  movel([-0.151447, -0.814996, -2.788348, -1.109046, 1.570796, 1.419350],accel_mss,speed_ms,0,blend_radius_m)
  movel([-0.155435, -0.823121, -2.786879, -1.102389, 1.570796, 1.415362],accel_mss,speed_ms,0,blend_radius_m)
  movel([-0.157149, -0.827095, -2.786148, -1.099146, 1.570796, 1.413648],accel_mss,speed_ms,0,blend_radius_m)
  movel([-0.159989, -0.834849, -2.784696, -1.092844, 1.570796, 1.410807],accel_mss,speed_ms,0,blend_radius_m)
  movel([-0.161109, -0.838634, -2.783975, -1.089780, 1.570796, 1.409688],accel_mss,speed_ms,0,blend_radius_m)
  movel([-0.162732, -0.846011, -2.782547, -1.083831, 1.570796, 1.408064],accel_mss,speed_ms,0,blend_radius_m)
  movel([-0.163230, -0.849609, -2.781839, -1.080941, 1.570796, 1.407566],accel_mss,speed_ms,0,blend_radius_m)
  movel([-0.163513, -0.853139, -2.781138, -1.078112, 1.570796, 1.407283],accel_mss,speed_ms,0,blend_radius_m)
  movel([-0.163602, -0.858015, -2.780157, -1.074217, 1.570796, 1.407194],accel_mss,speed_ms,0,blend_radius_m)
  movel([-0.163380, -0.862704, -2.779201, -1.070483, 1.570796, 1.407417],accel_mss,speed_ms,0,blend_radius_m)
  movel([-0.162870, -0.867194, -2.778274, -1.066921, 1.570796, 1.407926],accel_mss,speed_ms,0,blend_radius_m)
  movel([-0.162104, -0.871488, -2.777376, -1.063525, 1.570796, 1.408692],accel_mss,speed_ms,0,blend_radius_m)
  movel([-0.161097, -0.875560, -2.776515, -1.060315, 1.570796, 1.409700],accel_mss,speed_ms,0,blend_radius_m)
  movel([-0.159870, -0.879398, -2.775693, -1.057297, 1.570796, 1.410927],accel_mss,speed_ms,0,blend_radius_m)
  movel([-0.158448, -0.882999, -2.774915, -1.054475, 1.570796, 1.412348],accel_mss,speed_ms,0,blend_radius_m)
  movel([-0.156848, -0.886344, -2.774185, -1.051861, 1.570796, 1.413948],accel_mss,speed_ms,0,blend_radius_m)
  movel([-0.149158, -0.898055, -2.771574, -1.042759, 1.570796, 1.421638],accel_mss,speed_ms,0,blend_radius_m)
  movel([-0.143209, -0.907609, -2.769382, -1.035398, 1.570796, 1.427587],accel_mss,speed_ms,0,blend_radius_m)
  movel([-0.142775, -0.908633, -2.769143, -1.034613, 1.570796, 1.428021],accel_mss,speed_ms,0,blend_radius_m)
  movel([-0.135600, -0.899262, -2.771300, -1.041826, 1.570796, 1.435197],accel_mss,speed_ms,0,blend_radius_m)
  movel([-0.127938, -0.890014, -2.773376, -1.048999, 1.570796, 1.442859],accel_mss,speed_ms,0,blend_radius_m)
  movel([-0.119839, -0.880922, -2.775365, -1.056102, 1.570796, 1.450957],accel_mss,speed_ms,0,blend_radius_m)
  movel([-0.111369, -0.872030, -2.777262, -1.063097, 1.570796, 1.459427],accel_mss,speed_ms,0,blend_radius_m)
  movel([-0.102591, -0.863390, -2.779061, -1.069938, 1.570796, 1.468205],accel_mss,speed_ms,0,blend_radius_m)
  movel([-0.093574, -0.855040, -2.780757, -1.076592, 1.570796, 1.477222],accel_mss,speed_ms,0,blend_radius_m)
  movel([-0.084386, -0.847036, -2.782346, -1.083007, 1.570796, 1.486410],accel_mss,speed_ms,0,blend_radius_m)
  movel([-0.075105, -0.839424, -2.783823, -1.089142, 1.570796, 1.495692],accel_mss,speed_ms,0,blend_radius_m)
  movel([-0.070692, -0.836034, -2.784471, -1.091884, 1.570796, 1.500104],accel_mss,speed_ms,0,blend_radius_m)
  movel([-0.066171, -0.832804, -2.785082, -1.094503, 1.570796, 1.504626],accel_mss,speed_ms,0,blend_radius_m)
  movel([-0.061579, -0.829772, -2.785650, -1.096967, 1.570796, 1.509218],accel_mss,speed_ms,0,blend_radius_m)
  movel([-0.056967, -0.826981, -2.786169, -1.099239, 1.570796, 1.513830],accel_mss,speed_ms,0,blend_radius_m)
  movel([-0.052375, -0.824471, -2.786631, -1.101286, 1.570796, 1.518421],accel_mss,speed_ms,0,blend_radius_m)
  movel([-0.047846, -0.822284, -2.787032, -1.103074, 1.570796, 1.522951],accel_mss,speed_ms,0,blend_radius_m)
  movel([-0.043425, -0.820455, -2.787365, -1.104569, 1.570796, 1.527371],accel_mss,speed_ms,0,blend_radius_m)
  movel([-0.039161, -0.819026, -2.787624, -1.105740, 1.570796, 1.531636],accel_mss,speed_ms,0,blend_radius_m)
  movel([-0.035094, -0.818037, -2.787802, -1.106550, 1.570796, 1.535702],accel_mss,speed_ms,0,blend_radius_m)
  movel([-0.031268, -0.817523, -2.787894, -1.106971, 1.570796, 1.539528],accel_mss,speed_ms,0,blend_radius_m)
  movel([-0.027734, -0.817526, -2.787894, -1.106969, 1.570796, 1.543062],accel_mss,speed_ms,0,blend_radius_m)
  movel([-0.024533, -0.818078, -2.787795, -1.106516, 1.570796, 1.546264],accel_mss,speed_ms,0,blend_radius_m)
  movel([-0.021709, -0.819214, -2.787590, -1.105586, 1.570796, 1.549087],accel_mss,speed_ms,0,blend_radius_m)
  movel([-0.019297, -0.820962, -2.787273, -1.104155, 1.570796, 1.551499],accel_mss,speed_ms,0,blend_radius_m)
  movel([-0.017345, -0.823352, -2.786837, -1.102201, 1.570796, 1.553452],accel_mss,speed_ms,0,blend_radius_m)
  movel([-0.015891, -0.826416, -2.786273, -1.099700, 1.570796, 1.554905],accel_mss,speed_ms,0,blend_radius_m)
  movel([-0.014708, -0.831178, -2.785387, -1.095824, 1.570796, 1.556088],accel_mss,speed_ms,0,blend_radius_m)
  movel([-0.014174, -0.836590, -2.784365, -1.091434, 1.570796, 1.556622],accel_mss,speed_ms,0,blend_radius_m)
  movel([-0.014196, -0.842501, -2.783230, -1.086658, 1.570796, 1.556600],accel_mss,speed_ms,0,blend_radius_m)
  movel([-0.014673, -0.848767, -2.782005, -1.081616, 1.570796, 1.556123],accel_mss,speed_ms,0,blend_radius_m)
  movel([-0.015515, -0.855244, -2.780716, -1.076429, 1.570796, 1.555282],accel_mss,speed_ms,0,blend_radius_m)
  movel([-0.016634, -0.861800, -2.779387, -1.071202, 1.570796, 1.554162],accel_mss,speed_ms,0,blend_radius_m)
  movel([-0.019330, -0.874610, -2.776716, -1.061062, 1.570796, 1.551466],accel_mss,speed_ms,0,blend_radius_m)
  movel([-0.021385, -0.882738, -2.774972, -1.054680, 1.570796, 1.549411],accel_mss,speed_ms,0,blend_radius_m)
  movel([-0.023782, -0.890821, -2.773197, -1.048372, 1.570796, 1.547015],accel_mss,speed_ms,0,blend_radius_m)
  movel([-0.026474, -0.898860, -2.771392, -1.042138, 1.570796, 1.544323],accel_mss,speed_ms,0,blend_radius_m)
  movel([-0.029419, -0.906874, -2.769553, -1.035963, 1.570796, 1.541377],accel_mss,speed_ms,0,blend_radius_m)
  movel([-0.032573, -0.914860, -2.767679, -1.029850, 1.570796, 1.538223],accel_mss,speed_ms,0,blend_radius_m)
  movel([-0.035892, -0.922833, -2.765768, -1.023788, 1.570796, 1.534904],accel_mss,speed_ms,0,blend_radius_m)
  movel([-0.042880, -0.938782, -2.761820, -1.011787, 1.570796, 1.527916],accel_mss,speed_ms,0,blend_radius_m)
  movel([-0.036325, -0.939075, -2.761746, -1.011568, 1.570796, 1.534471],accel_mss,speed_ms,0,blend_radius_m)
  movel([-0.032953, -0.939481, -2.761643, -1.011265, 1.570796, 1.537843],accel_mss,speed_ms,0,blend_radius_m)
  movel([-0.030089, -0.940387, -2.761414, -1.010589, 1.570796, 1.540707],accel_mss,speed_ms,0,blend_radius_m)
  movel([-0.028984, -0.941104, -2.761231, -1.010053, 1.570796, 1.541813],accel_mss,speed_ms,0,blend_radius_m)
  movel([-0.028168, -0.942040, -2.760993, -1.009356, 1.570796, 1.542628],accel_mss,speed_ms,0,blend_radius_m)
  movel([-0.027690, -0.943217, -2.760692, -1.008479, 1.570796, 1.543106],accel_mss,speed_ms,0,blend_radius_m)
  movel([-0.027603, -0.944666, -2.760321, -1.007402, 1.570796, 1.543193],accel_mss,speed_ms,0,blend_radius_m)
  movel([-0.027958, -0.946409, -2.759872, -1.006107, 1.570796, 1.542838],accel_mss,speed_ms,0,blend_radius_m)
  movel([-0.028810, -0.948485, -2.759335, -1.004569, 1.570796, 1.541986],accel_mss,speed_ms,0,blend_radius_m)
  movel([-0.030204, -0.950916, -2.758703, -1.002770, 1.570796, 1.540592],accel_mss,speed_ms,0,blend_radius_m)
  movel([-0.032189, -0.953722, -2.757967, -1.000700, 1.570796, 1.538607],accel_mss,speed_ms,0,blend_radius_m)
  movel([-0.034030, -0.956006, -2.757365, -0.999018, 1.570796, 1.536766],accel_mss,speed_ms,0,blend_radius_m)
  movel([-0.035882, -0.958061, -2.756820, -0.997508, 1.570796, 1.534914],accel_mss,speed_ms,0,blend_radius_m)
  movel([-0.037742, -0.959903, -2.756328, -0.996157, 1.570796, 1.533055],accel_mss,speed_ms,0,blend_radius_m)
  movel([-0.041487, -0.963031, -2.755489, -0.993869, 1.570796, 1.529310],accel_mss,speed_ms,0,blend_radius_m)
  movel([-0.043369, -0.964351, -2.755133, -0.992905, 1.570796, 1.527427],accel_mss,speed_ms,0,blend_radius_m)
  movel([-0.047159, -0.966604, -2.754522, -0.991264, 1.570796, 1.523638],accel_mss,speed_ms,0,blend_radius_m)
  movel([-0.050963, -0.968447, -2.754019, -0.989923, 1.570796, 1.519833],accel_mss,speed_ms,0,blend_radius_m)
  movel([-0.054779, -0.970023, -2.753588, -0.988778, 1.570796, 1.516017],accel_mss,speed_ms,0,blend_radius_m)
  movel([-0.062394, -0.972906, -2.752793, -0.986690, 1.570796, 1.508402],accel_mss,speed_ms,0,blend_radius_m)
  movel([-0.066370, -0.979281, -2.751016, -0.982092, 1.570796, 1.504426],accel_mss,speed_ms,0,blend_radius_m)
  movel([-0.068546, -0.982465, -2.750118, -0.979807, 1.570796, 1.502250],accel_mss,speed_ms,0,blend_radius_m)
  movel([-0.070857, -0.985559, -2.749237, -0.977593, 1.570796, 1.499939],accel_mss,speed_ms,0,blend_radius_m)
  movel([-0.073309, -0.988496, -2.748395, -0.975498, 1.570796, 1.497488],accel_mss,speed_ms,0,blend_radius_m)
  movel([-0.075903, -0.991209, -2.747612, -0.973569, 1.570796, 1.494894],accel_mss,speed_ms,0,blend_radius_m)
  movel([-0.078648, -0.993632, -2.746907, -0.971850, 1.570796, 1.492149],accel_mss,speed_ms,0,blend_radius_m)
  movel([-0.081555, -0.995707, -2.746300, -0.970382, 1.570796, 1.489241],accel_mss,speed_ms,0,blend_radius_m)
  movel([-0.083598, -0.996753, -2.745993, -0.969643, 1.570796, 1.487198],accel_mss,speed_ms,0,blend_radius_m)
  movel([-0.085214, -0.997109, -2.745888, -0.969392, 1.570796, 1.485582],accel_mss,speed_ms,0,blend_radius_m)
  movel([-0.086450, -0.996877, -2.745957, -0.969556, 1.570796, 1.484347],accel_mss,speed_ms,0,blend_radius_m)
  movel([-0.087346, -0.996152, -2.746170, -0.970067, 1.570796, 1.483451],accel_mss,speed_ms,0,blend_radius_m)
  movel([-0.087946, -0.995031, -2.746498, -0.970860, 1.570796, 1.482851],accel_mss,speed_ms,0,blend_radius_m)
  movel([-0.088287, -0.993617, -2.746911, -0.971861, 1.570796, 1.482509],accel_mss,speed_ms,0,blend_radius_m)
  movel([-0.088418, -0.992006, -2.747380, -0.973003, 1.570796, 1.482378],accel_mss,speed_ms,0,blend_radius_m)
  movel([-0.088369, -0.990291, -2.747877, -0.974221, 1.570796, 1.482428],accel_mss,speed_ms,0,blend_radius_m)
  movel([-0.087893, -0.986486, -2.748972, -0.976931, 1.570796, 1.482904],accel_mss,speed_ms,0,blend_radius_m)
  movel([-0.087059, -0.982547, -2.750094, -0.979748, 1.570796, 1.483737],accel_mss,speed_ms,0,blend_radius_m)
  movel([-0.084858, -0.974333, -2.752398, -0.985658, 1.570796, 1.485939],accel_mss,speed_ms,0,blend_radius_m)
  movel([-0.093540, -0.972916, -2.752791, -0.986682, 1.570796, 1.477256],accel_mss,speed_ms,0,blend_radius_m)
  movel([-0.102455, -0.971877, -2.753077, -0.987434, 1.570796, 1.468341],accel_mss,speed_ms,0,blend_radius_m)
  movel([-0.111365, -0.970808, -2.753372, -0.988209, 1.570796, 1.459431],accel_mss,speed_ms,0,blend_radius_m)
  movel([-0.115747, -0.970134, -2.753557, -0.988698, 1.570796, 1.455049],accel_mss,speed_ms,0,blend_radius_m)
  movel([-0.120046, -0.969296, -2.753787, -0.989306, 1.570796, 1.450750],accel_mss,speed_ms,0,blend_radius_m)
  movel([-0.124039, -0.968285, -2.754064, -0.990041, 1.570796, 1.446757],accel_mss,speed_ms,0,blend_radius_m)
  movel([-0.127889, -0.967094, -2.754388, -0.990906, 1.570796, 1.442907],accel_mss,speed_ms,0,blend_radius_m)
  movel([-0.135327, -0.964371, -2.755127, -0.992891, 1.570796, 1.435469],accel_mss,speed_ms,0,blend_radius_m)
  movel([-0.142709, -0.961582, -2.755879, -0.994928, 1.570796, 1.428087],accel_mss,speed_ms,0,blend_radius_m)
  movel([-0.150371, -0.959179, -2.756522, -0.996688, 1.570796, 1.420425],accel_mss,speed_ms,0,blend_radius_m)
  movel([-0.152086, -0.963930, -2.755246, -0.993213, 1.570796, 1.418710],accel_mss,speed_ms,0,blend_radius_m)
  movel([-0.153549, -0.968557, -2.753989, -0.989843, 1.570796, 1.417247],accel_mss,speed_ms,0,blend_radius_m)
  movel([-0.154762, -0.973052, -2.752753, -0.986584, 1.570796, 1.416035],accel_mss,speed_ms,0,blend_radius_m)
  movel([-0.155729, -0.977408, -2.751541, -0.983440, 1.570796, 1.415067],accel_mss,speed_ms,0,blend_radius_m)
  movel([-0.156451, -0.981621, -2.750356, -0.980411, 1.570796, 1.414345],accel_mss,speed_ms,0,blend_radius_m)
  movel([-0.156938, -0.985687, -2.749200, -0.977501, 1.570796, 1.413859],accel_mss,speed_ms,0,blend_radius_m)
  movel([-0.157185, -0.989600, -2.748077, -0.974712, 1.570796, 1.413612],accel_mss,speed_ms,0,blend_radius_m)
  movel([-0.157205, -0.993359, -2.746986, -0.972043, 1.570796, 1.413592],accel_mss,speed_ms,0,blend_radius_m)
  movel([-0.156995, -0.996957, -2.745933, -0.969499, 1.570796, 1.413802],accel_mss,speed_ms,0,blend_radius_m)
  movel([-0.156554, -1.000385, -2.744920, -0.967083, 1.570796, 1.414242],accel_mss,speed_ms,0,blend_radius_m)
  movel([-0.155895, -1.003650, -2.743948, -0.964791, 1.570796, 1.414901],accel_mss,speed_ms,0,blend_radius_m)
  movel([-0.155018, -1.006740, -2.743020, -0.962629, 1.570796, 1.415778],accel_mss,speed_ms,0,blend_radius_m)
  movel([-0.153919, -1.009647, -2.742140, -0.960602, 1.570796, 1.416877],accel_mss,speed_ms,0,blend_radius_m)
  movel([-0.152607, -1.012377, -2.741308, -0.958704, 1.570796, 1.418189],accel_mss,speed_ms,0,blend_radius_m)
  movel([-0.151084, -1.014919, -2.740528, -0.956942, 1.570796, 1.419713],accel_mss,speed_ms,0,blend_radius_m)
  movel([-0.149346, -1.017271, -2.739802, -0.955317, 1.570796, 1.421450],accel_mss,speed_ms,0,blend_radius_m)
  movel([-0.146282, -1.020526, -2.738789, -0.953073, 1.570796, 1.424514],accel_mss,speed_ms,0,blend_radius_m)
  movel([-0.142850, -1.023308, -2.737918, -0.951163, 1.570796, 1.427946],accel_mss,speed_ms,0,blend_radius_m)
  movel([-0.139097, -1.025667, -2.737174, -0.949548, 1.570796, 1.431699],accel_mss,speed_ms,0,blend_radius_m)
  movel([-0.135055, -1.027644, -2.736547, -0.948198, 1.570796, 1.435741],accel_mss,speed_ms,0,blend_radius_m)
  movel([-0.130770, -1.029287, -2.736024, -0.947078, 1.570796, 1.440026],accel_mss,speed_ms,0,blend_radius_m)
  movel([-0.126280, -1.030634, -2.735593, -0.946162, 1.570796, 1.444516],accel_mss,speed_ms,0,blend_radius_m)
  movel([-0.121626, -1.031732, -2.735241, -0.945416, 1.570796, 1.449171],accel_mss,speed_ms,0,blend_radius_m)
  movel([-0.116838, -1.032609, -2.734959, -0.944821, 1.570796, 1.453958],accel_mss,speed_ms,0,blend_radius_m)
  movel([-0.106974, -1.033936, -2.734531, -0.943921, 1.570796, 1.463822],accel_mss,speed_ms,0,blend_radius_m)
  movel([-0.096981, -1.035022, -2.734180, -0.943187, 1.570796, 1.473815],accel_mss,speed_ms,0,blend_radius_m)
  movel([-0.089406, -1.036121, -2.733824, -0.942444, 1.570796, 1.481391],accel_mss,speed_ms,0,blend_radius_m)
  movel([-0.086797, -1.036293, -2.733768, -0.942328, 1.570796, 1.484000],accel_mss,speed_ms,0,blend_radius_m)
  movel([-0.082087, -1.036201, -2.733798, -0.942390, 1.570796, 1.488709],accel_mss,speed_ms,0,blend_radius_m)
  movel([-0.081105, -1.036377, -2.733741, -0.942271, 1.570796, 1.489692],accel_mss,speed_ms,0,blend_radius_m)
  movel([-0.080223, -1.036750, -2.733620, -0.942019, 1.570796, 1.490574],accel_mss,speed_ms,0,blend_radius_m)
  movel([-0.079458, -1.037384, -2.733413, -0.941592, 1.570796, 1.491338],accel_mss,speed_ms,0,blend_radius_m)
  movel([-0.078830, -1.038339, -2.733102, -0.940948, 1.570796, 1.491966],accel_mss,speed_ms,0,blend_radius_m)
  movel([-0.078371, -1.039682, -2.732663, -0.940044, 1.570796, 1.492426],accel_mss,speed_ms,0,blend_radius_m)
  movel([-0.078211, -1.041203, -2.732164, -0.939022, 1.570796, 1.492585],accel_mss,speed_ms,0,blend_radius_m)
  movel([-0.078322, -1.042870, -2.731615, -0.937905, 1.570796, 1.492474],accel_mss,speed_ms,0,blend_radius_m)
  movel([-0.078680, -1.044666, -2.731020, -0.936703, 1.570796, 1.492116],accel_mss,speed_ms,0,blend_radius_m)
  movel([-0.079260, -1.046558, -2.730392, -0.935440, 1.570796, 1.491536],accel_mss,speed_ms,0,blend_radius_m)
  movel([-0.080989, -1.050554, -2.729054, -0.932781, 1.570796, 1.489808],accel_mss,speed_ms,0,blend_radius_m)
  movel([-0.082090, -1.052608, -2.728361, -0.931420, 1.570796, 1.488706],accel_mss,speed_ms,0,blend_radius_m)
  movel([-0.084632, -1.056710, -2.726966, -0.928713, 1.570796, 1.486165],accel_mss,speed_ms,0,blend_radius_m)
  movel([-0.087485, -1.060661, -2.725610, -0.926118, 1.570796, 1.483311],accel_mss,speed_ms,0,blend_radius_m)
  movel([-0.090454, -1.064281, -2.724356, -0.923752, 1.570796, 1.480342],accel_mss,speed_ms,0,blend_radius_m)
  movel([-0.093367, -1.067405, -2.723264, -0.921720, 1.570796, 1.477429],accel_mss,speed_ms,0,blend_radius_m)
  movel([-0.097927, -1.071627, -2.721776, -0.918986, 1.570796, 1.472870],accel_mss,speed_ms,0,blend_radius_m)
  movel([-0.100289, -1.073583, -2.721081, -0.917725, 1.570796, 1.470507],accel_mss,speed_ms,0,blend_radius_m)
  movel([-0.102689, -1.075423, -2.720424, -0.916541, 1.570796, 1.468107],accel_mss,speed_ms,0,blend_radius_m)
  movel([-0.107574, -1.078758, -2.719227, -0.914404, 1.570796, 1.463222],accel_mss,speed_ms,0,blend_radius_m)
  movel([-0.112504, -1.081599, -2.718199, -0.912591, 1.570796, 1.458292],accel_mss,speed_ms,0,blend_radius_m)
  movel([-0.117406, -1.083911, -2.717357, -0.911121, 1.570796, 1.453391],accel_mss,speed_ms,0,blend_radius_m)
  movel([-0.122195, -1.085658, -2.716717, -0.910013, 1.570796, 1.448602],accel_mss,speed_ms,0,blend_radius_m)
  movel([-0.124527, -1.086307, -2.716479, -0.909603, 1.570796, 1.446270],accel_mss,speed_ms,0,blend_radius_m)
  movel([-0.129018, -1.087135, -2.716175, -0.909079, 1.570796, 1.441778],accel_mss,speed_ms,0,blend_radius_m)
  movel([-0.131158, -1.087301, -2.716114, -0.908974, 1.570796, 1.439638],accel_mss,speed_ms,0,blend_radius_m)
  movel([-0.133875, -1.087278, -2.716122, -0.908989, 1.570796, 1.436921],accel_mss,speed_ms,0,blend_radius_m)
  movel([-0.136457, -1.087013, -2.716220, -0.909156, 1.570796, 1.434339],accel_mss,speed_ms,0,blend_radius_m)
  movel([-0.138916, -1.086536, -2.716395, -0.909458, 1.570796, 1.431880],accel_mss,speed_ms,0,blend_radius_m)
  movel([-0.141274, -1.085885, -2.716634, -0.909870, 1.570796, 1.429522],accel_mss,speed_ms,0,blend_radius_m)
  movel([-0.145748, -1.084182, -2.717258, -0.910949, 1.570796, 1.425048],accel_mss,speed_ms,0,blend_radius_m)
  movel([-0.150009, -1.082170, -2.717991, -0.912228, 1.570796, 1.420787],accel_mss,speed_ms,0,blend_radius_m)
  movel([-0.155186, -1.079424, -2.718986, -0.913979, 1.570796, 1.415610],accel_mss,speed_ms,0,blend_radius_m)
  movel([-0.160187, -1.076374, -2.720084, -0.915931, 1.570796, 1.410610],accel_mss,speed_ms,0,blend_radius_m)
  movel([-0.164967, -1.072997, -2.721289, -0.918102, 1.570796, 1.405830],accel_mss,speed_ms,0,blend_radius_m)
  movel([-0.169489, -1.069278, -2.722606, -0.920505, 1.570796, 1.401308],accel_mss,speed_ms,0,blend_radius_m)
  movel([-0.173708, -1.065187, -2.724040, -0.923162, 1.570796, 1.397089],accel_mss,speed_ms,0,blend_radius_m)
  movel([-0.177576, -1.060702, -2.725596, -0.926091, 1.570796, 1.393221],accel_mss,speed_ms,0,blend_radius_m)
  movel([-0.181051, -1.055798, -2.727278, -0.929314, 1.570796, 1.389745],accel_mss,speed_ms,0,blend_radius_m)
  movel([-0.184087, -1.050445, -2.729090, -0.932854, 1.570796, 1.386710],accel_mss,speed_ms,0,blend_radius_m)
  movel([-0.186073, -1.046124, -2.730536, -0.935729, 1.570796, 1.384723],accel_mss,speed_ms,0,blend_radius_m)
  movel([-0.187880, -1.041406, -2.732097, -0.938886, 1.570796, 1.382916],accel_mss,speed_ms,0,blend_radius_m)
  movel([-0.189439, -1.036317, -2.733760, -0.942311, 1.570796, 1.381358],accel_mss,speed_ms,0,blend_radius_m)
  movel([-0.190682, -1.030894, -2.735510, -0.945985, 1.570796, 1.380114],accel_mss,speed_ms,0,blend_radius_m)
  movel([-0.191534, -1.025166, -2.737332, -0.949891, 1.570796, 1.379263],accel_mss,speed_ms,0,blend_radius_m)
  movel([-0.191918, -1.019165, -2.739214, -0.954010, 1.570796, 1.378878],accel_mss,speed_ms,0,blend_radius_m)
  movel([-0.191763, -1.012919, -2.741142, -0.958328, 1.570796, 1.379033],accel_mss,speed_ms,0,blend_radius_m)
  movel([-0.191455, -1.009712, -2.742120, -0.960557, 1.570796, 1.379341],accel_mss,speed_ms,0,blend_radius_m)
  movel([-0.190983, -1.006458, -2.743105, -0.962827, 1.570796, 1.379813],accel_mss,speed_ms,0,blend_radius_m)
  movel([-0.189719, -1.000183, -2.744980, -0.967225, 1.570796, 1.381077],accel_mss,speed_ms,0,blend_radius_m)
  movel([-0.188031, -0.993695, -2.746888, -0.971805, 1.570796, 1.382765],accel_mss,speed_ms,0,blend_radius_m)
  movel([-0.185918, -0.987014, -2.748821, -0.976555, 1.570796, 1.384878],accel_mss,speed_ms,0,blend_radius_m)
  movel([-0.183392, -0.980165, -2.750768, -0.981457, 1.570796, 1.387404],accel_mss,speed_ms,0,blend_radius_m)
  movel([-0.180442, -0.973167, -2.752721, -0.986500, 1.570796, 1.390354],accel_mss,speed_ms,0,blend_radius_m)
  movel([-0.177085, -0.966055, -2.754671, -0.991663, 1.570796, 1.393711],accel_mss,speed_ms,0,blend_radius_m)
  movel([-0.173317, -0.958850, -2.756610, -0.996929, 1.570796, 1.397479],accel_mss,speed_ms,0,blend_radius_m)
  movel([-0.169142, -0.951585, -2.758528, -1.002276, 1.570796, 1.401654],accel_mss,speed_ms,0,blend_radius_m)
  movel([-0.177984, -0.943954, -2.760504, -1.007931, 1.570796, 1.392812],accel_mss,speed_ms,0,blend_radius_m)
  movel([-0.182461, -0.940170, -2.761469, -1.010750, 1.570796, 1.388335],accel_mss,speed_ms,0,blend_radius_m)
  movel([-0.186722, -0.936099, -2.762496, -1.013794, 1.570796, 1.384074],accel_mss,speed_ms,0,blend_radius_m)
  movel([-0.189559, -0.932656, -2.763356, -1.016376, 1.570796, 1.381237],accel_mss,speed_ms,0,blend_radius_m)
  movel([-0.191976, -0.928741, -2.764325, -1.019323, 1.570796, 1.378820],accel_mss,speed_ms,0,blend_radius_m)
  movel([-0.193988, -0.924385, -2.765391, -1.022612, 1.570796, 1.376808],accel_mss,speed_ms,0,blend_radius_m)
  movel([-0.195602, -0.919608, -2.766546, -1.026235, 1.570796, 1.375194],accel_mss,speed_ms,0,blend_radius_m)
  movel([-0.196828, -0.914436, -2.767780, -1.030173, 1.570796, 1.373968],accel_mss,speed_ms,0,blend_radius_m)
  movel([-0.197671, -0.908892, -2.769083, -1.034414, 1.570796, 1.373125],accel_mss,speed_ms,0,blend_radius_m)
  movel([-0.198141, -0.902999, -2.770447, -1.038943, 1.570796, 1.372655],accel_mss,speed_ms,0,blend_radius_m)
  movel([-0.198246, -0.896786, -2.771861, -1.043741, 1.570796, 1.372550],accel_mss,speed_ms,0,blend_radius_m)
  movel([-0.197990, -0.890280, -2.773317, -1.048792, 1.570796, 1.372806],accel_mss,speed_ms,0,blend_radius_m)
  movel([-0.197379, -0.883499, -2.774806, -1.054084, 1.570796, 1.373418],accel_mss,speed_ms,0,blend_radius_m)
  movel([-0.196419, -0.876474, -2.776320, -1.059595, 1.570796, 1.374377],accel_mss,speed_ms,0,blend_radius_m)
  movel([-0.195120, -0.869237, -2.777848, -1.065304, 1.570796, 1.375676],accel_mss,speed_ms,0,blend_radius_m)
  movel([-0.193486, -0.861813, -2.779384, -1.071192, 1.570796, 1.377310],accel_mss,speed_ms,0,blend_radius_m)
  movel([-0.191530, -0.854245, -2.780917, -1.077227, 1.570796, 1.379267],accel_mss,speed_ms,0,blend_radius_m)
  movel([-0.189249, -0.846551, -2.782441, -1.083397, 1.570796, 1.381547],accel_mss,speed_ms,0,blend_radius_m)
  movel([-0.186663, -0.838776, -2.783948, -1.089666, 1.570796, 1.384133],accel_mss,speed_ms,0,blend_radius_m)
  movel([-0.181160, -0.823879, -2.786740, -1.101770, 1.570796, 1.389637],accel_mss,speed_ms,0,blend_radius_m)
  movel([-0.178053, -0.816218, -2.788129, -1.108042, 1.570796, 1.392744],accel_mss,speed_ms,0,blend_radius_m)
  movel([-0.174652, -0.808422, -2.789510, -1.114457, 1.570796, 1.396144],accel_mss,speed_ms,0,blend_radius_m)
  movel([-0.170903, -0.800498, -2.790880, -1.121010, 1.570796, 1.399893],accel_mss,speed_ms,0,blend_radius_m)
  movel([-0.166766, -0.792462, -2.792237, -1.127690, 1.570796, 1.404030],accel_mss,speed_ms,0,blend_radius_m)
  movel([-0.162191, -0.784317, -2.793578, -1.134494, 1.570796, 1.408605],accel_mss,speed_ms,0,blend_radius_m)
  movel([-0.157128, -0.776076, -2.794900, -1.141412, 1.570796, 1.413668],accel_mss,speed_ms,0,blend_radius_m)
  movel([-0.150973, -0.766860, -2.796339, -1.149190, 1.570796, 1.419823],accel_mss,speed_ms,0,blend_radius_m)
  movel([-0.144342, -0.757619, -2.797739, -1.157031, 1.570796, 1.426454],accel_mss,speed_ms,0,blend_radius_m)
  movel([-0.137271, -0.748380, -2.799097, -1.164911, 1.570796, 1.433525],accel_mss,speed_ms,0,blend_radius_m)
  movel([-0.129792, -0.739184, -2.800409, -1.172797, 1.570796, 1.441004],accel_mss,speed_ms,0,blend_radius_m)
  movel([-0.121944, -0.730069, -2.801669, -1.180651, 1.570796, 1.448852],accel_mss,speed_ms,0,blend_radius_m)
  movel([-0.113770, -0.721080, -2.802874, -1.188435, 1.570796, 1.457026],accel_mss,speed_ms,0,blend_radius_m)
  movel([-0.105305, -0.712251, -2.804022, -1.196116, 1.570796, 1.465492],accel_mss,speed_ms,0,blend_radius_m)
  movel([-0.096600, -0.703635, -2.805107, -1.203647, 1.570796, 1.474197],accel_mss,speed_ms,0,blend_radius_m)
  movel([-0.087699, -0.695278, -2.806128, -1.210982, 1.570796, 1.483097],accel_mss,speed_ms,0,blend_radius_m)
  movel([-0.078662, -0.687228, -2.807083, -1.218079, 1.570796, 1.492134],accel_mss,speed_ms,0,blend_radius_m)
  movel([-0.069532, -0.679533, -2.807968, -1.224888, 1.570796, 1.501264],accel_mss,speed_ms,0,blend_radius_m)
  movel([-0.060365, -0.672240, -2.808784, -1.231364, 1.570796, 1.510431],accel_mss,speed_ms,0,blend_radius_m)
  movel([-0.051227, -0.665407, -2.809528, -1.237454, 1.570796, 1.519569],accel_mss,speed_ms,0,blend_radius_m)
  movel([-0.042167, -0.659076, -2.810199, -1.243114, 1.570796, 1.528629],accel_mss,speed_ms,0,blend_radius_m)
  movel([-0.033247, -0.653297, -2.810797, -1.248295, 1.570796, 1.537549],accel_mss,speed_ms,0,blend_radius_m)
  movel([-0.024524, -0.648122, -2.811321, -1.252946, 1.570796, 1.546273],accel_mss,speed_ms,0,blend_radius_m)
  movel([-0.015396, -0.643113, -2.811817, -1.257459, 1.570796, 1.555400],accel_mss,speed_ms,0,blend_radius_m)
  movel([-0.006368, -0.638517, -2.812264, -1.261608, 1.570796, 1.564428],accel_mss,speed_ms,0,blend_radius_m)
  movel([0.002483, -0.634467, -2.812650, -1.265272, 1.570796, 1.573279],accel_mss,speed_ms,0,blend_radius_m)
  movel([0.011077, -0.631111, -2.812965, -1.268314, 1.570796, 1.581874],accel_mss,speed_ms,0,blend_radius_m)
  movel([0.020717, -0.628189, -2.813235, -1.270964, 1.570796, 1.591514],accel_mss,speed_ms,0,blend_radius_m)
  movel([0.029958, -0.626311, -2.813407, -1.272670, 1.570796, 1.600754],accel_mss,speed_ms,0,blend_radius_m)
  movel([0.038695, -0.625494, -2.813481, -1.273413, 1.570796, 1.609491],accel_mss,speed_ms,0,blend_radius_m)
  movel([0.046827, -0.625746, -2.813459, -1.273184, 1.570796, 1.617623],accel_mss,speed_ms,0,blend_radius_m)
  movel([0.054267, -0.627064, -2.813338, -1.271987, 1.570796, 1.625063],accel_mss,speed_ms,0,blend_radius_m)
  movel([0.060928, -0.629437, -2.813120, -1.269832, 1.570796, 1.631725],accel_mss,speed_ms,0,blend_radius_m)
  movel([0.066738, -0.632841, -2.812803, -1.266745, 1.570796, 1.637535],accel_mss,speed_ms,0,blend_radius_m)
  movel([0.071630, -0.637250, -2.812385, -1.262754, 1.570796, 1.642427],accel_mss,speed_ms,0,blend_radius_m)
  movel([0.080139, -0.647263, -2.811407, -1.253719, 1.570796, 1.650935],accel_mss,speed_ms,0,blend_radius_m)
  movel([0.083892, -0.652766, -2.810852, -1.248771, 1.570796, 1.654688],accel_mss,speed_ms,0,blend_radius_m)
  movel([0.087126, -0.658973, -2.810210, -1.243206, 1.570796, 1.657922],accel_mss,speed_ms,0,blend_radius_m)
  movel([0.092254, -0.669756, -2.809057, -1.233576, 1.570796, 1.663050],accel_mss,speed_ms,0,blend_radius_m)
  movel([0.095202, -0.674825, -2.808498, -1.229066, 1.570796, 1.665998],accel_mss,speed_ms,0,blend_radius_m)
  movel([0.098521, -0.679457, -2.807977, -1.224955, 1.570796, 1.669318],accel_mss,speed_ms,0,blend_radius_m)
  movel([0.102318, -0.683483, -2.807517, -1.221389, 1.570796, 1.673114],accel_mss,speed_ms,0,blend_radius_m)
  movel([0.106666, -0.686745, -2.807139, -1.218505, 1.570796, 1.677463],accel_mss,speed_ms,0,blend_radius_m)
  movel([0.111676, -0.689079, -2.806866, -1.216444, 1.570796, 1.682472],accel_mss,speed_ms,0,blend_radius_m)
  movel([0.117434, -0.690323, -2.806719, -1.215347, 1.570796, 1.688231],accel_mss,speed_ms,0,blend_radius_m)
  movel([0.120030, -0.690376, -2.806713, -1.215300, 1.570796, 1.690827],accel_mss,speed_ms,0,blend_radius_m)
  movel([0.122938, -0.689845, -2.806775, -1.215768, 1.570796, 1.693735],accel_mss,speed_ms,0,blend_radius_m)
  movel([0.124501, -0.689269, -2.806843, -1.216277, 1.570796, 1.695297],accel_mss,speed_ms,0,blend_radius_m)
  movel([0.126126, -0.688444, -2.806940, -1.217005, 1.570796, 1.696922],accel_mss,speed_ms,0,blend_radius_m)
  movel([0.127815, -0.687331, -2.807071, -1.217988, 1.570796, 1.698611],accel_mss,speed_ms,0,blend_radius_m)
  movel([0.129555, -0.685891, -2.807238, -1.219259, 1.570796, 1.700351],accel_mss,speed_ms,0,blend_radius_m)
  movel([0.131319, -0.684125, -2.807443, -1.220821, 1.570796, 1.702115],accel_mss,speed_ms,0,blend_radius_m)
  movel([0.132980, -0.682166, -2.807668, -1.222555, 1.570796, 1.703776],accel_mss,speed_ms,0,blend_radius_m)
  movel([0.135970, -0.677934, -2.808149, -1.226306, 1.570796, 1.706767],accel_mss,speed_ms,0,blend_radius_m)
  movel([0.137783, -0.674917, -2.808487, -1.228985, 1.570796, 1.708580],accel_mss,speed_ms,0,blend_radius_m)
  movel([0.139361, -0.671936, -2.808818, -1.231635, 1.570796, 1.710157],accel_mss,speed_ms,0,blend_radius_m)
  movel([0.141870, -0.666110, -2.809452, -1.236827, 1.570796, 1.712666],accel_mss,speed_ms,0,blend_radius_m)
  movel([0.143598, -0.660509, -2.810049, -1.241832, 1.570796, 1.714394],accel_mss,speed_ms,0,blend_radius_m)
  movel([0.144658, -0.655168, -2.810605, -1.246616, 1.570796, 1.715454],accel_mss,speed_ms,0,blend_radius_m)
  movel([0.145152, -0.650148, -2.811117, -1.251123, 1.570796, 1.715948],accel_mss,speed_ms,0,blend_radius_m)
  movel([0.145192, -0.645490, -2.811583, -1.255316, 1.570796, 1.715988],accel_mss,speed_ms,0,blend_radius_m)
  movel([0.144887, -0.641239, -2.812000, -1.259149, 1.570796, 1.715683],accel_mss,speed_ms,0,blend_radius_m)
  movel([0.143440, -0.633449, -2.812746, -1.266194, 1.570796, 1.714237],accel_mss,speed_ms,0,blend_radius_m)
  movel([0.142144, -0.629825, -2.813084, -1.269480, 1.570796, 1.712941],accel_mss,speed_ms,0,blend_radius_m)
  movel([0.140471, -0.626589, -2.813382, -1.272418, 1.570796, 1.711267],accel_mss,speed_ms,0,blend_radius_m)
  movel([0.138417, -0.623775, -2.813637, -1.274977, 1.570796, 1.709214],accel_mss,speed_ms,0,blend_radius_m)
  movel([0.135985, -0.621398, -2.813850, -1.277141, 1.570796, 1.706781],accel_mss,speed_ms,0,blend_radius_m)
  movel([0.133177, -0.619487, -2.814020, -1.278882, 1.570796, 1.703974],accel_mss,speed_ms,0,blend_radius_m)
  movel([0.130010, -0.618050, -2.814147, -1.280192, 1.570796, 1.700806],accel_mss,speed_ms,0,blend_radius_m)
  movel([0.126480, -0.617113, -2.814229, -1.281047, 1.570796, 1.697276],accel_mss,speed_ms,0,blend_radius_m)
  speed_ms = 0.005
  movel([0.126480, -0.611489, -2.807428, -1.293472, 1.570796, 1.697276],accel_mss,speed_ms,0,blend_radius_m)
  speed_ms = 0.040
  movel([0.123325, -0.648612, -2.803909, -1.259867, 1.570796, 1.694121],accel_mss,speed_ms,0,blend_radius_m)
  speed_ms = 0.005
  movel([0.123325, -0.654823, -2.810641, -1.246925, 1.570796, 1.694121],accel_mss,speed_ms,0,blend_radius_m)
  speed_ms = 0.025
  movel([0.118895, -0.654079, -2.810717, -1.247593, 1.570796, 1.689691],accel_mss,speed_ms,0,blend_radius_m)
  movel([0.113905, -0.654220, -2.810703, -1.247466, 1.570796, 1.684701],accel_mss,speed_ms,0,blend_radius_m)
  movel([0.111148, -0.654809, -2.810642, -1.246938, 1.570796, 1.681944],accel_mss,speed_ms,0,blend_radius_m)
  movel([0.108196, -0.655839, -2.810536, -1.246014, 1.570796, 1.678993],accel_mss,speed_ms,0,blend_radius_m)
  movel([0.105036, -0.657380, -2.810376, -1.244633, 1.570796, 1.675833],accel_mss,speed_ms,0,blend_radius_m)
  movel([0.101649, -0.659496, -2.810155, -1.242737, 1.570796, 1.672446],accel_mss,speed_ms,0,blend_radius_m)
  speed_ms = 0.005
  movel([0.101649, -0.653216, -2.803433, -1.255740, 1.570796, 1.672446],accel_mss,speed_ms,0,blend_radius_m)
  speed_ms = 0.040
  movel([0.112275, -0.638238, -2.804950, -1.269201, 1.570796, 1.683072],accel_mss,speed_ms,0,blend_radius_m)
  speed_ms = 0.005
  movel([0.112275, -0.644289, -2.811702, -1.256398, 1.570796, 1.683072],accel_mss,speed_ms,0,blend_radius_m)
  speed_ms = 0.025
  movel([0.112399, -0.639470, -2.812172, -1.260747, 1.570796, 1.683195],accel_mss,speed_ms,0,blend_radius_m)
  movel([0.111517, -0.635629, -2.812540, -1.264220, 1.570796, 1.682314],accel_mss,speed_ms,0,blend_radius_m)
  movel([0.109701, -0.632797, -2.812807, -1.266785, 1.570796, 1.680497],accel_mss,speed_ms,0,blend_radius_m)
  movel([0.107011, -0.631035, -2.812972, -1.268382, 1.570796, 1.677807],accel_mss,speed_ms,0,blend_radius_m)
  movel([0.103521, -0.630378, -2.813033, -1.268978, 1.570796, 1.674318],accel_mss,speed_ms,0,blend_radius_m)
  movel([0.099319, -0.630861, -2.812988, -1.268540, 1.570796, 1.670115],accel_mss,speed_ms,0,blend_radius_m)
  movel([0.094491, -0.632506, -2.812834, -1.267049, 1.570796, 1.665287],accel_mss,speed_ms,0,blend_radius_m)
  movel([0.091867, -0.633776, -2.812715, -1.265898, 1.570796, 1.662663],accel_mss,speed_ms,0,blend_radius_m)
  movel([0.089124, -0.635335, -2.812568, -1.264486, 1.570796, 1.659920],accel_mss,speed_ms,0,blend_radius_m)
  speed_ms = 0.005
  movel([0.089124, -0.629423, -2.805799, -1.277167, 1.570796, 1.659920],accel_mss,speed_ms,0,blend_radius_m)
  speed_ms = 0.040
  movel([0.102652, -0.614078, -2.807201, -1.291111, 1.570796, 1.673448],accel_mss,speed_ms,0,blend_radius_m)
  speed_ms = 0.005
  movel([0.102652, -0.619744, -2.813997, -1.278647, 1.570796, 1.673448],accel_mss,speed_ms,0,blend_radius_m)
  speed_ms = 0.025
  movel([0.102279, -0.617703, -2.814177, -1.280509, 1.570796, 1.673075],accel_mss,speed_ms,0,blend_radius_m)
  movel([0.101580, -0.615933, -2.814332, -1.282124, 1.570796, 1.672376],accel_mss,speed_ms,0,blend_radius_m)
  movel([0.099284, -0.613217, -2.814567, -1.284605, 1.570796, 1.670080],accel_mss,speed_ms,0,blend_radius_m)
  movel([0.095934, -0.611616, -2.814704, -1.286069, 1.570796, 1.666730],accel_mss,speed_ms,0,blend_radius_m)
  movel([0.091712, -0.611145, -2.814744, -1.286500, 1.570796, 1.662509],accel_mss,speed_ms,0,blend_radius_m)
  movel([0.086803, -0.611795, -2.814689, -1.285905, 1.570796, 1.657599],accel_mss,speed_ms,0,blend_radius_m)
  movel([0.081418, -0.613547, -2.814538, -1.284303, 1.570796, 1.652214],accel_mss,speed_ms,0,blend_radius_m)
  movel([0.078603, -0.614838, -2.814427, -1.283124, 1.570796, 1.649399],accel_mss,speed_ms,0,blend_radius_m)
  movel([0.072873, -0.618207, -2.814133, -1.280049, 1.570796, 1.643669],accel_mss,speed_ms,0,blend_radius_m)
  movel([0.070007, -0.620280, -2.813950, -1.278159, 1.570796, 1.640803],accel_mss,speed_ms,0,blend_radius_m)
  speed_ms = 0.005
  movel([0.070007, -0.614605, -2.807154, -1.290630, 1.570796, 1.640803],accel_mss,speed_ms,0,blend_radius_m)
  speed_ms = 0.040
  movel([0.089300, -0.594878, -2.808821, -1.308690, 1.570796, 1.660097],accel_mss,speed_ms,0,blend_radius_m)
  speed_ms = 0.005
  movel([0.089300, -0.600228, -2.815650, -1.296511, 1.570796, 1.660097],accel_mss,speed_ms,0,blend_radius_m)
  speed_ms = 0.025
  movel([0.085848, -0.598031, -2.815827, -1.298531, 1.570796, 1.656644],accel_mss,speed_ms,0,blend_radius_m)
  movel([0.081583, -0.596921, -2.815915, -1.299553, 1.570796, 1.652379],accel_mss,speed_ms,0,blend_radius_m)
  movel([0.076593, -0.596959, -2.815912, -1.299518, 1.570796, 1.647389],accel_mss,speed_ms,0,blend_radius_m)
  movel([0.070948, -0.598187, -2.815814, -1.298388, 1.570796, 1.641744],accel_mss,speed_ms,0,blend_radius_m)
  movel([0.064745, -0.600651, -2.815616, -1.296122, 1.570796, 1.635541],accel_mss,speed_ms,0,blend_radius_m)
  movel([0.061464, -0.602352, -2.815477, -1.294559, 1.570796, 1.632260],accel_mss,speed_ms,0,blend_radius_m)
  movel([0.058084, -0.604371, -2.815312, -1.292707, 1.570796, 1.628881],accel_mss,speed_ms,0,blend_radius_m)
  movel([0.054609, -0.606713, -2.815118, -1.290558, 1.570796, 1.625405],accel_mss,speed_ms,0,blend_radius_m)
  movel([0.051053, -0.609382, -2.814894, -1.288113, 1.570796, 1.621849],accel_mss,speed_ms,0,blend_radius_m)
  movel([0.047438, -0.612369, -2.814640, -1.285380, 1.570796, 1.618234],accel_mss,speed_ms,0,blend_radius_m)
  movel([0.043773, -0.615680, -2.814354, -1.282355, 1.570796, 1.614569],accel_mss,speed_ms,0,blend_radius_m)
  speed_ms = 0.005
  movel([0.043773, -0.610078, -2.807551, -1.294760, 1.570796, 1.614569],accel_mss,speed_ms,0,blend_radius_m)
  speed_ms = 0.040
  movel([0.064233, -0.586313, -2.809497, -1.316579, 1.570796, 1.635029],accel_mss,speed_ms,0,blend_radius_m)
  speed_ms = 0.005
  movel([0.064233, -0.591518, -2.816339, -1.304531, 1.570796, 1.635029],accel_mss,speed_ms,0,blend_radius_m)
  speed_ms = 0.025
  movel([0.063094, -0.589044, -2.816530, -1.306816, 1.570796, 1.633890],accel_mss,speed_ms,0,blend_radius_m)
  movel([0.061364, -0.587230, -2.816668, -1.308492, 1.570796, 1.632160],accel_mss,speed_ms,0,blend_radius_m)
  movel([0.059073, -0.586116, -2.816752, -1.309521, 1.570796, 1.629869],accel_mss,speed_ms,0,blend_radius_m)
  movel([0.056266, -0.585735, -2.816781, -1.309874, 1.570796, 1.627062],accel_mss,speed_ms,0,blend_radius_m)
  movel([0.052290, -0.586217, -2.816744, -1.309427, 1.570796, 1.623086],accel_mss,speed_ms,0,blend_radius_m)
  movel([0.047869, -0.587504, -2.816647, -1.308238, 1.570796, 1.618665],accel_mss,speed_ms,0,blend_radius_m)
  movel([0.042312, -0.589762, -2.816475, -1.306152, 1.570796, 1.613109],accel_mss,speed_ms,0,blend_radius_m)
  movel([0.036448, -0.592816, -2.816238, -1.303335, 1.570796, 1.607244],accel_mss,speed_ms,0,blend_radius_m)
  movel([0.030360, -0.596687, -2.815934, -1.299768, 1.570796, 1.601157],accel_mss,speed_ms,0,blend_radius_m)
  movel([0.024131, -0.601411, -2.815554, -1.295424, 1.570796, 1.594927],accel_mss,speed_ms,0,blend_radius_m)
  movel([0.017873, -0.606995, -2.815094, -1.290300, 1.570796, 1.588669],accel_mss,speed_ms,0,blend_radius_m)
  movel([0.014803, -0.610065, -2.814836, -1.287488, 1.570796, 1.585600],accel_mss,speed_ms,0,blend_radius_m)
  movel([0.008947, -0.616633, -2.814271, -1.281485, 1.570796, 1.579743],accel_mss,speed_ms,0,blend_radius_m)
  movel([0.006216, -0.620075, -2.813968, -1.278346, 1.570796, 1.577013],accel_mss,speed_ms,0,blend_radius_m)
  movel([0.003666, -0.623589, -2.813654, -1.275146, 1.570796, 1.574462],accel_mss,speed_ms,0,blend_radius_m)
  movel([0.001318, -0.627153, -2.813330, -1.271906, 1.570796, 1.572114],accel_mss,speed_ms,0,blend_radius_m)
  speed_ms = 0.005
  movel([0.001318, -0.621369, -2.806547, -1.284473, 1.570796, 1.572114],accel_mss,speed_ms,0,blend_radius_m)
  speed_ms = 0.040
  movel([0.022676, -0.589066, -2.809283, -1.314040, 1.570796, 1.593472],accel_mss,speed_ms,0,blend_radius_m)
  speed_ms = 0.005
  movel([0.022676, -0.594318, -2.816121, -1.301950, 1.570796, 1.593472],accel_mss,speed_ms,0,blend_radius_m)
  speed_ms = 0.025
  movel([0.015376, -0.597704, -2.815853, -1.298833, 1.570796, 1.586173],accel_mss,speed_ms,0,blend_radius_m)
  movel([0.007626, -0.602096, -2.815498, -1.294794, 1.570796, 1.578423],accel_mss,speed_ms,0,blend_radius_m)
  movel([-0.000368, -0.607465, -2.815055, -1.289870, 1.570796, 1.570428],accel_mss,speed_ms,0,blend_radius_m)
  movel([-0.004391, -0.610495, -2.814799, -1.287095, 1.570796, 1.566405],accel_mss,speed_ms,0,blend_radius_m)
  movel([-0.008399, -0.613754, -2.814521, -1.284114, 1.570796, 1.562398],accel_mss,speed_ms,0,blend_radius_m)
  movel([-0.012357, -0.617227, -2.814219, -1.280943, 1.570796, 1.558439],accel_mss,speed_ms,0,blend_radius_m)
  movel([-0.016240, -0.620904, -2.813894, -1.277591, 1.570796, 1.554557],accel_mss,speed_ms,0,blend_radius_m)
  movel([-0.020025, -0.624783, -2.813546, -1.274060, 1.570796, 1.550771],accel_mss,speed_ms,0,blend_radius_m)
  movel([-0.023687, -0.628860, -2.813173, -1.270356, 1.570796, 1.547109],accel_mss,speed_ms,0,blend_radius_m)
  movel([-0.027206, -0.633124, -2.812776, -1.266489, 1.570796, 1.543591],accel_mss,speed_ms,0,blend_radius_m)
  movel([-0.030543, -0.637564, -2.812355, -1.262470, 1.570796, 1.540253],accel_mss,speed_ms,0,blend_radius_m)
  movel([-0.033686, -0.642176, -2.811909, -1.258304, 1.570796, 1.537111],accel_mss,speed_ms,0,blend_radius_m)
  movel([-0.036604, -0.646954, -2.811438, -1.253997, 1.570796, 1.534193],accel_mss,speed_ms,0,blend_radius_m)
  speed_ms = 0.005
  movel([-0.036604, -0.640863, -2.804691, -1.266835, 1.570796, 1.534193],accel_mss,speed_ms,0,blend_radius_m)
  speed_ms = 0.040
  movel([-0.022149, -0.609169, -2.807629, -1.295591, 1.570796, 1.548647],accel_mss,speed_ms,0,blend_radius_m)
  speed_ms = 0.005
  movel([-0.022149, -0.614755, -2.814434, -1.283200, 1.570796, 1.548647],accel_mss,speed_ms,0,blend_radius_m)
  speed_ms = 0.025
  movel([-0.025873, -0.616783, -2.814258, -1.281348, 1.570796, 1.544923],accel_mss,speed_ms,0,blend_radius_m)
  movel([-0.029708, -0.619203, -2.814045, -1.279141, 1.570796, 1.541089],accel_mss,speed_ms,0,blend_radius_m)
  movel([-0.033605, -0.621987, -2.813798, -1.276604, 1.570796, 1.537191],accel_mss,speed_ms,0,blend_radius_m)
  movel([-0.037532, -0.625097, -2.813518, -1.273774, 1.570796, 1.533264],accel_mss,speed_ms,0,blend_radius_m)
  movel([-0.041453, -0.628505, -2.813206, -1.270678, 1.570796, 1.529343],accel_mss,speed_ms,0,blend_radius_m)
  movel([-0.045324, -0.632175, -2.812865, -1.267348, 1.570796, 1.525473],accel_mss,speed_ms,0,blend_radius_m)
  movel([-0.049105, -0.636067, -2.812498, -1.263824, 1.570796, 1.521691],accel_mss,speed_ms,0,blend_radius_m)
  movel([-0.052772, -0.640159, -2.812105, -1.260125, 1.570796, 1.518024],accel_mss,speed_ms,0,blend_radius_m)
  movel([-0.056275, -0.644407, -2.811690, -1.256292, 1.570796, 1.514522],accel_mss,speed_ms,0,blend_radius_m)
  movel([-0.059585, -0.648764, -2.811257, -1.252368, 1.570796, 1.511211],accel_mss,speed_ms,0,blend_radius_m)
  movel([-0.062677, -0.653185, -2.810809, -1.248396, 1.570796, 1.508120],accel_mss,speed_ms,0,blend_radius_m)
  movel([-0.065528, -0.657633, -2.810350, -1.244406, 1.570796, 1.505269],accel_mss,speed_ms,0,blend_radius_m)
  movel([-0.068119, -0.662068, -2.809884, -1.240437, 1.570796, 1.502677],accel_mss,speed_ms,0,blend_radius_m)
  movel([-0.070432, -0.666459, -2.809415, -1.236515, 1.570796, 1.500365],accel_mss,speed_ms,0,blend_radius_m)
  movel([-0.072431, -0.670752, -2.808948, -1.232689, 1.570796, 1.498365],accel_mss,speed_ms,0,blend_radius_m)
  movel([-0.074111, -0.674922, -2.808487, -1.228980, 1.570796, 1.496685],accel_mss,speed_ms,0,blend_radius_m)
  speed_ms = 0.005
  movel([-0.074111, -0.668415, -2.801797, -1.242177, 1.570796, 1.496685],accel_mss,speed_ms,0,blend_radius_m)
  speed_ms = 0.040
  movel([-0.066858, -0.641711, -2.804607, -1.266071, 1.570796, 1.503938],accel_mss,speed_ms,0,blend_radius_m)
  speed_ms = 0.005
  movel([-0.066858, -0.647816, -2.811352, -1.253221, 1.570796, 1.503938],accel_mss,speed_ms,0,blend_radius_m)
  speed_ms = 0.025
  movel([-0.070442, -0.650003, -2.811132, -1.251254, 1.570796, 1.500354],accel_mss,speed_ms,0,blend_radius_m)
  movel([-0.074094, -0.652775, -2.810851, -1.248763, 1.570796, 1.496702],accel_mss,speed_ms,0,blend_radius_m)
  movel([-0.077748, -0.656034, -2.810516, -1.245839, 1.570796, 1.493049],accel_mss,speed_ms,0,blend_radius_m)
  movel([-0.081363, -0.659683, -2.810136, -1.242571, 1.570796, 1.489434],accel_mss,speed_ms,0,blend_radius_m)
  movel([-0.084887, -0.663631, -2.809718, -1.239040, 1.570796, 1.485909],accel_mss,speed_ms,0,blend_radius_m)
  movel([-0.088268, -0.667779, -2.809272, -1.235338, 1.570796, 1.482528],accel_mss,speed_ms,0,blend_radius_m)
  movel([-0.091469, -0.672036, -2.808807, -1.231546, 1.570796, 1.479327],accel_mss,speed_ms,0,blend_radius_m)
  movel([-0.094435, -0.676312, -2.808332, -1.227745, 1.570796, 1.476361],accel_mss,speed_ms,0,blend_radius_m)
  movel([-0.097268, -0.680725, -2.807833, -1.223832, 1.570796, 1.473529],accel_mss,speed_ms,0,blend_radius_m)
  movel([-0.099872, -0.685149, -2.807325, -1.219916, 1.570796, 1.470924],accel_mss,speed_ms,0,blend_radius_m)
  movel([-0.102209, -0.689533, -2.806812, -1.216044, 1.570796, 1.468587],accel_mss,speed_ms,0,blend_radius_m)
  movel([-0.104211, -0.693806, -2.806305, -1.212278, 1.570796, 1.466585],accel_mss,speed_ms,0,blend_radius_m)
  movel([-0.105837, -0.697907, -2.805810, -1.208672, 1.570796, 1.464959],accel_mss,speed_ms,0,blend_radius_m)
  movel([-0.107039, -0.701777, -2.805337, -1.205275, 1.570796, 1.463757],accel_mss,speed_ms,0,blend_radius_m)
  movel([-0.107755, -0.705352, -2.804893, -1.202143, 1.570796, 1.463041],accel_mss,speed_ms,0,blend_radius_m)
  movel([-0.107950, -0.708578, -2.804488, -1.199322, 1.570796, 1.462846],accel_mss,speed_ms,0,blend_radius_m)
  speed_ms = 0.005
  movel([-0.107950, -0.701603, -2.797873, -1.212913, 1.570796, 1.462846],accel_mss,speed_ms,0,blend_radius_m)
  speed_ms = 0.040
  movel([-0.110320, -0.684454, -2.799961, -1.227974, 1.570796, 1.460476],accel_mss,speed_ms,0,blend_radius_m)
  speed_ms = 0.005
  movel([-0.110320, -0.691191, -2.806616, -1.214581, 1.570796, 1.460476],accel_mss,speed_ms,0,blend_radius_m)
  speed_ms = 0.025
  movel([-0.115088, -0.696403, -2.805993, -1.209993, 1.570796, 1.455708],accel_mss,speed_ms,0,blend_radius_m)
  movel([-0.119860, -0.702223, -2.805282, -1.204884, 1.570796, 1.450936],accel_mss,speed_ms,0,blend_radius_m)
  movel([-0.124369, -0.708375, -2.804514, -1.199500, 1.570796, 1.446427],accel_mss,speed_ms,0,blend_radius_m)
  movel([-0.128353, -0.714586, -2.803722, -1.194082, 1.570796, 1.442443],accel_mss,speed_ms,0,blend_radius_m)
  movel([-0.131570, -0.720601, -2.802937, -1.188851, 1.570796, 1.439226],accel_mss,speed_ms,0,blend_radius_m)
  movel([-0.132817, -0.723461, -2.802559, -1.186369, 1.570796, 1.437979],accel_mss,speed_ms,0,blend_radius_m)
  movel([-0.133780, -0.726174, -2.802196, -1.184019, 1.570796, 1.437016],accel_mss,speed_ms,0,blend_radius_m)
  movel([-0.134435, -0.728723, -2.801852, -1.181814, 1.570796, 1.436361],accel_mss,speed_ms,0,blend_radius_m)
  movel([-0.134755, -0.731074, -2.801532, -1.179782, 1.570796, 1.436041],accel_mss,speed_ms,0,blend_radius_m)
  movel([-0.134702, -0.733189, -2.801242, -1.177958, 1.570796, 1.436094],accel_mss,speed_ms,0,blend_radius_m)
  movel([-0.134258, -0.735056, -2.800984, -1.176348, 1.570796, 1.436538],accel_mss,speed_ms,0,blend_radius_m)
  speed_ms = 0.005
  movel([-0.134258, -0.727738, -2.794433, -1.190218, 1.570796, 1.436538],accel_mss,speed_ms,0,blend_radius_m)
  speed_ms = 0.040
  movel([-0.143177, -0.726739, -2.794570, -1.191080, 1.570796, 1.427620],accel_mss,speed_ms,0,blend_radius_m)
  speed_ms = 0.005
  movel([-0.143177, -0.734045, -2.801124, -1.177220, 1.570796, 1.427620],accel_mss,speed_ms,0,blend_radius_m)
  speed_ms = 0.025
  movel([-0.148309, -0.742676, -2.799916, -1.169798, 1.570796, 1.422487],accel_mss,speed_ms,0,blend_radius_m)
  movel([-0.150599, -0.746995, -2.799297, -1.166096, 1.570796, 1.420197],accel_mss,speed_ms,0,blend_radius_m)
  movel([-0.152589, -0.751214, -2.798685, -1.162489, 1.570796, 1.418207],accel_mss,speed_ms,0,blend_radius_m)
  movel([-0.154194, -0.755273, -2.798088, -1.159028, 1.570796, 1.416602],accel_mss,speed_ms,0,blend_radius_m)
  movel([-0.155337, -0.759108, -2.797516, -1.155765, 1.570796, 1.415460],accel_mss,speed_ms,0,blend_radius_m)
  movel([-0.155927, -0.762648, -2.796982, -1.152759, 1.570796, 1.414869],accel_mss,speed_ms,0,blend_radius_m)
  movel([-0.155895, -0.765842, -2.796495, -1.150052, 1.570796, 1.414902],accel_mss,speed_ms,0,blend_radius_m)
  speed_ms = 0.005
  # Splitting Linear movement in 2 (instruction 3386: MoveL 3110)
  movel([-0.155895, -0.747318, -2.780284, -1.184788, 1.570796, 1.414902],accel_mss,speed_ms,0,blend_radius_m)
  movel([-0.155895, -0.730984, -2.763964, -1.217440, 1.570796, 1.414902],accel_mss,speed_ms,0,blend_radius_m)
  speed_ms = 1.000
  movel([-0.155895, -0.730984, -2.763964, -1.217440, 1.570796, 1.414902],accel_mss,speed_ms,0,blend_radius_m)
  # Splitting Linear movement in 6 (instruction 3389: MoveL 3112)
  movel([-0.155895, -0.707995, -2.736548, -1.267846, 1.570796, 1.414902],accel_mss,speed_ms,0,blend_radius_m)
  movel([-0.155895, -0.689517, -2.708886, -1.313986, 1.570796, 1.414902],accel_mss,speed_ms,0,blend_radius_m)
  movel([-0.155895, -0.674819, -2.681001, -1.356569, 1.570796, 1.414902],accel_mss,speed_ms,0,blend_radius_m)
  movel([-0.155895, -0.663318, -2.652909, -1.396162, 1.570796, 1.414902],accel_mss,speed_ms,0,blend_radius_m)
  movel([-0.155895, -0.654540, -2.624621, -1.433227, 1.570796, 1.414902],accel_mss,speed_ms,0,blend_radius_m)
  movel([-0.155895, -0.648105, -2.596144, -1.468140, 1.570796, 1.414902],accel_mss,speed_ms,0,blend_radius_m)
  # End of main program
end

Machining1()
